(* IEC 61131-3 sources: kns-port-domestic/targets/astra/lib/src/POUs/Util/F_TimeToSec, 1 file *)

(* ---- F_TimeToSec.decl.st ---- *)
// Назначение: длительность TIME (мс) в секундах LREAL. TIME_TO_LREAL переводит 32-битное число
//             миллисекунд в LREAL точно.
// Автор:      kr0nsch
// Версия:     0.1.0
// Документ:   docs/fb/Functions.md
FUNCTION F_TimeToSec : LREAL
VAR_INPUT
    tIn : TIME;   // длительность
END_VAR
